(* IEC 61131-3 sources: cds-text-sync-reference-project/project-view/CODESYS_HMI/PLC Logic/HMI_Application/MFL_VISU, 3 files *)

(* ---- DUT_CONV_FRAME.st ---- *)
TYPE DUT_CONV_FRAME :
STRUCT
	conv_idx : INT := 1;      // Index in ZONE_MFL.g_aConfigs (1..4)
	sName : STRING(16);       // Safe name copy
	state : STRING(15);       // String representation of state
	//config : DUT_MFL_Config;  // Config copy for visualization
	dimension : INT := 50;    // [mm] segment size for ASCII
	pec_idx : USINT := 1;     // Which PEC to show slip for (1..10)
	iInstantSlip : INT;       // Current/Last measured slip [mm]

	// Compatibility fields for older Visu
	conv_number : INT;
	pec_choice : INT;
	pecAverageSlip : INT;

	asciiString : STRING(255); // The visual representation
END_STRUCT
END_TYPE

(* ---- ENUM_SegmentStatus.st ---- *)
{attribute 'qualified_only'}
{attribute 'strict'}
TYPE ENUM_SegmentStatus :
(
	Empty_Segment := 95,     // '_' Empty 50mm space
	Cargo_Start := 91,       // '[' Left boundary of cargo item
	Cargo_End := 93,         // ']' Right boundary of cargo item
	Cargo_Filled := 35,      // '#' Segment fully occupied by cargo
	Sensor_Inactive := 111,  // 'o' Sensor position, no cargo detected
	Sensor_Active := 120,    // 'x' Sensor position, cargo detected
	Conveyor_Start := 123,   // '{'  Start edge of conveyor
	Conveyor_End := 125,     // '}' end edge of conveyor
	NULL := 0				 // String termination
)USINT;
END_TYPE

(* ---- ZONE_HMI.st ---- *)
{attribute 'qualified_only'}
VAR_GLOBAL
    // === Global Commands (HMI -> PLC) ===
    xStart: BOOL; // Master Start pulse for all zones
    xStop: BOOL; // Master Stop pulse for all zones
    xReset: BOOL; // Master Reset for all errors
    xReverse: BOOL; // Global direction control (Logic Level)
    xEmitt1: BOOL;
    xEmitt2: BOOL;

    // === Global Status (PLC -> HMI) ===
    xAnyError: BOOL; // True if any zone in error state
    xAnyWarning: BOOL; // True if any zone has a warning
    xSystemOK: BOOL; // True if communication and all zones are OK
    xRunning: BOOL; // True if at least one conveyor is moving

    // === Visualization Mapping ===
    // This array holds references to the frames used by the HMI.
    // It is initialized in MAIN.st to point to VISUALIZATION.aFrames.
    arConveyors: ARRAY[1..4] OF DUT_CONV_FRAME;

	arErrors : ARRAY[0..10] OF BOOL;

END_VAR
